// TIA Portal V21 export
// export: Created 2026-11-11T00:48:31.540486Z, ExportSetting WithDefaults, DisplayName Totally Integrated Automation Portal, DisplayVersion V21 Update 3, DisplayName STEP 7 Professional, DisplayVersion V21 Update 3, DisplayName STEP 7 Safety, DisplayVersion V21, DisplayName Tech WebApplication, DisplayVersion V21, DisplayName WinCC Basic/Comfort/Advanced, DisplayVersion V21 Update 3, DisplayName WinCC Unified, DisplayVersion V21 Update 3
FUNCTION_BLOCK "FX_Fbd_160"   // FB238, FBD
{ S7_Optimized_Access := 'TRUE' }
VERSION : 0.1
// stored: AutoNumber true, IsIECCheckEnabled false, IsRetainMemResEnabled false, MemoryReserve 100, SetENOAutomatically false, UDAEnableTagReadback false
   VAR_INPUT
      "a" : Bool;
      "b" : Bool;
      c : Bool;
      ia : Int;
      ib : Int;
      ic : Int;
      da : DInt;
      db : DInt;
      ra : Real;
      rb : Real;
      wa : Word;
      wb : Word;
      dwa : DWord;
      ba : Byte;
      ta : Time;
      tb : Time;
      s1 : String;
      s2 : String;
   END_VAR
   VAR_OUTPUT
      q : Bool;
      q2 : Bool;
      io : Int;
      io2 : Int;
      dout : DInt;
      rout : Real;
      wout : Word;
      dwout : DWord;
      bout : Byte;
      tout : Time;
      sout : String;
   END_VAR
   VAR_IN_OUT
      arr : Array[0..9] of Int;
      barr : Array[0..7] of Bool;
      iinout : Int;
   END_VAR
   VAR
      inst : DRUM;
      ton1 { S7_SetPoint := 'True'} : TON_TIME;
      tof1 { S7_SetPoint := 'True'} : TOF_TIME;
      tp1 { S7_SetPoint := 'True'} : TP_TIME;
      tonr1 { S7_SetPoint := 'True'} : TONR_TIME;
      ctu1 { S7_SetPoint := 'True'} : CTU_INT;
      ctd1 { S7_SetPoint := 'True'} : CTD_INT;
      ctud1 { S7_SetPoint := 'True'} : CTUD_INT;
      rtrig1 { S7_SetPoint := 'True'} : R_TRIG;
      ftrig1 { S7_SetPoint := 'True'} : F_TRIG;
      edge1 : Bool;
      edge2 : Bool;
      stat1 : Bool;
      stat2 : Bool;
      stati : Int;
   END_VAR
   VAR_TEMP
      t1 : Bool;
      t2 : Bool;
      ti : Int;
      td : DInt;
      tr : Real;
      tw : Word;
      tt : Time;
      var1 : Variant;
   END_VAR
BEGIN

REGION Network 1: ---| |--- - Normally open contact
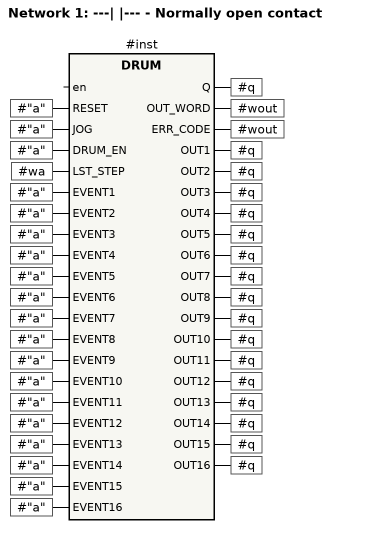
   #inst(RESET := #"a",   // DRUM
         JOG := #"a",
         DRUM_EN := #"a",
         LST_STEP := #wa,
         EVENT1 := #"a",
         EVENT2 := #"a",
         EVENT3 := #"a",
         EVENT4 := #"a",
         EVENT5 := #"a",
         EVENT6 := #"a",
         EVENT7 := #"a",
         EVENT8 := #"a",
         EVENT9 := #"a",
         EVENT10 := #"a",
         EVENT11 := #"a",
         EVENT12 := #"a",
         EVENT13 := #"a",
         EVENT14 := #"a",
         EVENT15 := #"a",
         EVENT16 := #"a",
         Q => #q,
         OUT_WORD => #wout,
         ERR_CODE => #wout,
         OUT1 => #q,
         OUT2 => #q,
         OUT3 => #q,
         OUT4 => #q,
         OUT5 => #q,
         OUT6 => #q,
         OUT7 => #q,
         OUT8 => #q,
         OUT9 => #q,
         OUT10 => #q,
         OUT11 => #q,
         OUT12 => #q,
         OUT13 => #q,
         OUT14 => #q,
         OUT15 => #q,
         OUT16 => #q);
END_REGION
END_FUNCTION_BLOCK
